// TIA Portal V21 export
// export: Created 2026-11-21T10:55:49.9625481Z, ExportSetting WithDefaults, DisplayName Totally Integrated Automation Portal, DisplayVersion V21, DisplayName STEP 7 Professional, DisplayVersion V21, DisplayName STEP 7 Safety, DisplayVersion V21, DisplayName Tech WebApplication, DisplayVersion V21, DisplayName WinCC Basic/Comfort/Advanced, DisplayVersion V21, DisplayName WinCC Unified, DisplayVersion V21
VAR_GLOBAL   // PLC tag table "IO"
   Run_North AT %I0.0 : Bool;   // Start the north station
   Lamp_North AT %Q0.0 : Bool;   // The north station runs
END_VAR
